// TIA Portal V21 export
// export: Created 2026-11-08T21:35:18.1521381Z, ExportSetting WithDefaults, DisplayName Totally Integrated Automation Portal, DisplayVersion V21 Update 3, DisplayName STEP 7 Professional, DisplayVersion V21 Update 3, DisplayName STEP 7 Safety, DisplayVersion V21, DisplayName Tech WebApplication, DisplayVersion V21, DisplayName WinCC Basic/Comfort/Advanced, DisplayVersion V21 Update 3, DisplayName WinCC Unified, DisplayVersion V21 Update 3
FUNCTION_BLOCK "FB_StlC_008"   // FB88, STL
TITLE = STL call PRESET_TIMER
{ S7_Optimized_Access := 'TRUE' }
VERSION : 0.1
// stored: AutoNumber true, IsRetainMemResEnabled false, MemoryReserve 100, UDAEnableTagReadback false
   VAR
      t1 { S7_SetPoint := 'True'} : IEC_TIMER;
   END_VAR
BEGIN

NETWORK
TITLE = 008 PRESET_TIMER
      CALL  PRESET_TIMER
      ( PT      := T#2S,
        "TIMER" := #t1
      );
END_FUNCTION_BLOCK
